Fanuc KAREL source: kd00040.KL

-- PROVISIONAL review KL for V940-1; original PC SHA256 de3c2b075bb72caab54953423af79fc80bc91ea5d329cbd03fa428a837b413b9
-- Incomplete behavior may be omitted. Consult companion uncertainty JSON. Do not deploy.
PROGRAM KD00040
%NOLOCKGROUP
BEGIN
  -- V9_ZERO_TABLE_METADATA_HINT layout=0001; no indexed target words; source/name/runtime held
  -- UNRESOLVED_PC offsets 5-26; opcodes AD,32,22,9B,9B,9C,9C,37,2C
  -- UNRESOLVED_PC offsets 31-35; opcodes 7F
END KD00040
